(* IEC 61131-3 sources: Test-Git_ESME26/TestProgettoESME_26.fbsproj/TemplateFullProgrammingFramework_Migration.device.xml.v3^/Plc Logic.plclogic.xml.v3^/Application.application.xml.v3^/TemplateFullProgrammingFramework/EquipmentModules/SR_CharlyModule.pou.xml.v3^, 9 files *)

(* ---- Init_Reactions.act.st ---- *)
__METADATA__
{
  "v3Meta": {
    "objectGuid": "4aa47ba2-99d8-49fa-95b1-7f556ffac844",
    "objectTypeGuid": "8ac092e5-3128-4e26-9e7e-11016c6684f2",
    "embeddedObjectTypeGuids": [
      "3b83b776-fb25-43b8-99f2-3c507c9143fc"
    ],
    "properties": {},
    "subObjects": {}
  }
}

(* System generated code, only to be changed by experienced programmers *)
IF c_udiNumberOfSubModules < 1 THEN
	RETURN;
END_IF

(* Change of default reactions only on demand *)
(* Compare SR MainMachine Action Init_Reactions *)

xInitReactionsException := FALSE;

(*****************************************************************************************************************************************************)
(* Init ReactionTranslationMode *)

TPL.FC_InitReactionTranslationMode(	i_udiNumberOfSubModules			:= c_udiNumberOfSubModules,
									i_petReactionTranslationMode	:= ADR(aetReactionTranslationMode),
									q_etDiag						=> etDiag,
									q_etDiagExt						=> etDiagExtTPL);

IF etDiag <> GD.ET_Diag.Ok AND NOT xInitReactionsException THEN
	xInitReactionsException := TRUE;

	stInitReactionsException.sMsg := SE_CTBX.FC_MultiConcat(i_sString1 := 'InitReactionTranslationMode - ',
														i_sString2 := GD.FC_EtDiagToString(i_etDiag := etDiag),
														i_sString3 := ' - ',
														i_sString4 := TPL.FC_EtDiagExtToString(i_etDiagExt := etDiagExtTPL));
END_IF

(*****************************************************************************************************************************************************)
(* Init ReactionTranslationTable *)

TPL.FC_InitReactionTranslationTable(i_udiNumberOfSubModules			:= c_udiNumberOfSubModules,
									i_pstReactionTranslationTable	:= ADR(aastReactionTranslationTable),
									q_etDiag						=> etDiag,
									q_etDiagExt						=> etDiagExtTPL);

IF etDiag <> GD.ET_Diag.Ok AND NOT xInitReactionsException THEN
	xInitReactionsException := TRUE;

	stInitReactionsException.sMsg := SE_CTBX.FC_MultiConcat(i_sString1 := 'InitReactionTranslationTable - ',
														i_sString2 := GD.FC_EtDiagToString(i_etDiag := etDiag),
														i_sString3 := ' - ',
														i_sString4 := TPL.FC_EtDiagExtToString(i_etDiagExt := etDiagExtTPL));
END_IF

(*****************************************************************************************************************************************************)
(* Init ReactionTranslationJobs *)

TPL.FC_InitReactionTranslationJobs( i_udiNumberOfSubModules			:= c_udiNumberOfSubModules,
									i_pstReactionTranslationJobs	:= ADR(astReactionTranslationJobs),
									q_etDiag						=> etDiag,
									q_etDiagExt						=> etDiagExtTPL);

IF etDiag <> GD.ET_Diag.Ok AND NOT xInitReactionsException THEN
	xInitReactionsException := TRUE;

	stInitReactionsException.sMsg := SE_CTBX.FC_MultiConcat(i_sString1 := 'InitReactionTranslationJobs - ',
														i_sString2 := GD.FC_EtDiagToString(i_etDiag := etDiag),
														i_sString3 := ' - ',
														i_sString4 := TPL.FC_EtDiagExtToString(i_etDiagExt := etDiagExtTPL));
END_IF

(*****************************************************************************************************************************************************)
(* Set exception if any exception occurred *)

fbExceptionHandler.SetException(i_xExceptionActive	:= xInitReactionsException,
								iq_stException		:= stInitReactionsException,
								iq_stExceptionList	:= iq_stExceptionList);

xInitSuccessful := xInitSuccessful AND NOT xInitReactionsException;

etDiag := GD.ET_Diag.Ok;
(* End of system generated code, only to be changed by experienced programmers *)

(* ---- Init_Slave3.act.st ---- *)
__METADATA__
{
  "v3Meta": {
    "objectGuid": "d2282e85-0a4e-4bdb-8c08-0233ce9aa560",
    "objectTypeGuid": "8ac092e5-3128-4e26-9e7e-11016c6684f2",
    "embeddedObjectTypeGuids": [
      "3b83b776-fb25-43b8-99f2-3c507c9143fc"
    ],
    "properties": {},
    "subObjects": {}
  }
}

(* System generated code, could be modified for your application *)

(* Standard interface *)
astSubModuleInterface[c_udiSlave3].i_sModuleName := CONCAT(STR1 := iq_stStandardModuleItf.i_sModuleName, STR2 := ': Slave3');

astSubModuleInterface[c_udiSlave3].i_xLogEnable     := TRUE;
astSubModuleInterface[c_udiSlave3].i_wLogDataFilter := UDINT_TO_WORD(TPL.ET_LogDataFilter.ModuleDefault);

fbSlave3Module.RegisterLoggerPoint(i_ifParent := fbLoggerPoint, i_sName := 'Slave3', q_etDiag :=, q_etDiagExt :=);

(* AxisModule specific interface *)
stSlave3Interface.stMain.i_ifMaster 		:= i_ifMaster; (* Master *)
stSlave3Interface.stMain.i_ifDrive  		:= DRV_Slave3.Axis;
stSlave3Interface.stMain.iq_lencEncoder		:= LE_Slave3.Axis;
DRV_Slave3.Axis.SetErrorStopRamp(i_lrDeceleration := 50_000,
								  i_lrJerk		  := 500_000);

xDriveIsVirtual := FC_IsDriveVirtual(	i_ifDrive	:= stSlave3Interface.stMain.i_ifDrive,
										q_etDiag	=> etDiag,
										q_etDiagExt	=> etDiagExt,
										q_sMsg		=> sMsgBuffer);

IF etDiag <> GD.ET_Diag.Ok AND NOT xIsDriveVirtualException THEN
	stIsDriveVirtualException.etDiag 	:= etDiag;
	stIsDriveVirtualException.udiDiagExt:= etDiagExt;
	stIsDriveVirtualException.sDiagExt 	:= FC_EtDiagExtToString(i_etDiagExt := etDiagExt);
	stIsDriveVirtualException.sMsg 		:= sMsgBuffer;
	xIsDriveVirtualException 			:= TRUE;
END_IF

fbExceptionHandler.SetException(i_xExceptionActive	:= xIsDriveVirtualException,
								iq_stException		:= stIsDriveVirtualException,
								iq_stExceptionList	:= iq_stExceptionList);

xInitSuccessful := xInitSuccessful AND NOT xIsDriveVirtualException;
etDiag := GD.ET_Diag.Ok;

stSlave3Interface.stMain.i_lrMotionActiveVelLimit := 15.0; (* Limit for max. velocity of astAxisModuleInterface to switch output AxisMove in Units/s *)
stSlave3Interface.stMain.i_etMotionActiveVelType  := AXM_ET_MotionActiveVelType.RefVelocity;

stSlave3Interface.stMain.i_timMasterStop := T#1S;
stSlave3Interface.stMain.i_xHwLimitPos   := FALSE;
stSlave3Interface.stMain.i_xHwLimitNeg   := FALSE;

stSlave3Interface.stMain.stReducedVelocity.i_xEnableReducedVelocity		:= FALSE;
stSlave3Interface.stMain.stReducedVelocity.i_xOnlyLimitCheck			:= FALSE;
stSlave3Interface.stMain.stReducedVelocity.i_lrMaxReducedVelocity		:= 50.0;

stSlave3Interface.stMain.i_xStart := FALSE;

(***************************************************************************************************************************************************************************************************)
(*** Homing ***)
	IF xDriveIsVirtual THEN
		stSlave3Interface.stHome.i_etMode := PDL_ET_HomeMode.SetPosAxisAndLogEncoderPosition;			(* Homing Mode  in case of virtual axis *)
	ELSE
		stSlave3Interface.stHome.i_etMode := PDL_ET_HomeMode.PosDirectionPosEdgeSensor;						(* Homing Mode in case of real axis *)
	END_IF

	stSlave3Interface.stHome.i_xEnableInitAbsReadPos := FALSE;		(* TRUE : Restores the AxisPosition depending on the stHome.etMode
																			  If stHome.i_etMode is equal to PDL_ET_HomeMode.RestorePosFromAxisEncoder or
																			  to PDL_ET_HomeMode.WriteAxisEncoder, the encoder of the axis is read,
																			  or else the position will be restored from the retain area *)

 	stSlave3Interface.stHome.stSetpos.iq_pstRestorePosRetain := ADR(Grp_stRestorePositionAxis4);

	stSlave3Interface.stHome.i_xResetHomeOk := FALSE;

	(* Possible modes for homing mode Sensor:
		PDL_ET_HomeMode.PosDirectionPosEdgeSensor
		PDL_ET_HomeMode.NegDirectionPosEdgeSensor
		PDL_ET_HomeMode.NegDirectionNegEdgeSensor
		PDL_ET_HomeMode.PosDirectionNegEdgeSensor
	*)
	stSlave3Interface.stHome.stSensor.i_lrHomePosition			:= 0.0;			(* Position at the end of homing in units *)
	stSlave3Interface.stHome.stSensor.i_lrVel					:= 10.0;		(* Homing ceiling velocity in units/s *)
	stSlave3Interface.stHome.stSensor.i_lrAcc					:= 1000.0;		(* Homing acceleration in units/s^2 *)
	stSlave3Interface.stHome.stSensor.i_lrDec					:= 1000.0;		(* Homing deceleration in units/s^2 *)
	stSlave3Interface.stHome.stSensor.i_lrJerk					:= 10000.0;		(* Homing jerk in units/s^3 *)
	stSlave3Interface.stHome.stSensor.i_lrOffset				:= 0.0;			(* Offset from home signal in units *)
	stSlave3Interface.stHome.stSensor.i_lrMaxTravel				:= 720.0;		(* Max. travel for referencing by normal input *)
	stSlave3Interface.stHome.stSensor.i_xRotativeSystem			:= FALSE;		(* Rotative system true or false for referencing by normal input *)
	stSlave3Interface.stHome.stSensor.i_xSensor					:= FALSE;		(* Input for home signal. Can be a signal from a controller input. Has to be written cyclic. *)

	(* Possible Modes for homing mode LimitSwitch:
		PDL_ET_HomeMode.PosDirectionPosEdgeHWLimitPos		normally open contact / Closing contact
		PDL_ET_HomeMode.NegDirectionPosEdgeHWLimitNeg		normally open contact / Closing contact
		PDL_ET_HomeMode.NegDirectionNegEdgeHWLimitNeg		normally closed contact / Opening contact
		PDL_ET_HomeMode.PosDirectionNegEdgeHWLimitPos		normally closed contact / Opening contact
	*)
	stSlave3Interface.stHome.stLimitSwitch.i_lrHomePosition		:= 0.0;			(* Position at the end of homing in units *)
	stSlave3Interface.stHome.stLimitSwitch.i_lrVel				:= 10.0;		(* Homing ceiling velocity in units/s *)
	stSlave3Interface.stHome.stLimitSwitch.i_lrLowVel			:= 5.0;			(* Homing low ceiling velocity in units/s *)
	stSlave3Interface.stHome.stLimitSwitch.i_lrAcc				:= 1000.0;		(* Homing acceleration in units/s^2 *)
	stSlave3Interface.stHome.stLimitSwitch.i_lrDec				:= 1000.0;		(* Homing deceleration in units/s^2 *)
	stSlave3Interface.stHome.stLimitSwitch.i_lrJerk				:= 10000.0;		(* Homing jerk in units/s^3 *)
	stSlave3Interface.stHome.stLimitSwitch.i_lrOffset			:= 0.0;			(* Offset from home signal in units *)
	stSlave3Interface.stHome.stLimitSwitch.i_lrMaxTravel		:= 9999.0;		(* Max. travel for referencing normal input as a hardware limit *)

	(* Possible modes for homing mode MoveOnPos:
		PDL_ET_HomeMode.MoveOnPosAbs
	*)
	stSlave3Interface.stHome.stMoveOnPos.i_lrTarget				:= 0.0;			(* Position at the end of homing in units *)
	stSlave3Interface.stHome.stMoveOnPos.i_lrVel				:= 10.0;		(* Homing ceiling velocity in units/s *)
	stSlave3Interface.stHome.stMoveOnPos.i_lrAcc				:= 1000.0;		(* Homing acceleration in units/s^2 *)
	stSlave3Interface.stHome.stMoveOnPos.i_lrDec				:= 1000.0;		(* Homing deceleration in units/s^2 *)
	stSlave3Interface.stHome.stMoveOnPos.i_lrJerk				:= 10000.0;		(* Homing jerk in units/s^3 *)
	stSlave3Interface.stHome.stMoveOnPos.i_lrPeriod				:= 0.0;			(* Period of the axis *)
	stSlave3Interface.stHome.stMoveOnPos.i_xRotativeSystem		:= FALSE;		(* Rotative system true or false *)

	(* Possible modes for homing mode SetPos:
		PDL_ET_HomeMode.SetPosAxisPosition
		PDL_ET_HomeMode.SetPosLogEncoderPosition
		PDL_ET_HomeMode.SetPosAxisAndLogEncoderPosition
		PDL_ET_HomeMode.RestorePosFromAxisEncoder
		PDL_ET_HomeMode.RestorePosFromRetain
	*)
	stSlave3Interface.stHome.stSetpos.i_lrHomePosition			:= 0.0;			(* Position at the end of homing in units *)
	stSlave3Interface.stHome.stSetpos.i_lrEncoderPosition		:= 0.0;			(* Encoder position in units after homing *)
	stSlave3Interface.stHome.stSetpos.i_lrAbsEncOffset			:= 100.0;		(* Distance to the jump of axis encoder in units  *)
	stSlave3Interface.stHome.stSetpos.i_lrRestoreWindow			:= 180;			(* How far can the drive be away from is correct position *)
	stSlave3Interface.stHome.stSetpos.i_lrUserPeriod			:= 360;			(* Period of the axis *)
	stSlave3Interface.stHome.stSetPos.i_xKeepPowerDisabled 		:= FALSE;		(* Keep Power disabled during SetPosHoming true or false*)

	(* Possible modes for homing mode Torque:
		PDL_ET_HomeMode.PosDirectionMaxTorque
		PDL_ET_HomeMode.NegDirectionMaxTorque
	*)
	stSlave3Interface.stHome.stTorque.i_lrHomePosition			:= 0.0;			(* Position at the end of homing in units *)
	stSlave3Interface.stHome.stTorque.i_lrVel					:= 10.0;		(* Homing ceiling velocity in units/s *)
	stSlave3Interface.stHome.stTorque.i_lrAcc					:= 1000.0;		(* Homing acceleration in units/s^2 *)
	stSlave3Interface.stHome.stTorque.i_lrDec					:= 1000.0;		(* Homing deceleration in units/s^2 *)
	stSlave3Interface.stHome.stTorque.i_lrJerk					:= 10000.0;		(* Homing jerk in units/s^3 *)
	stSlave3Interface.stHome.stTorque.i_lrOffset				:= 0.0;			(* Offset from home signal in units *)
	stSlave3Interface.stHome.stTorque.i_lrMaxTravel				:= 9999.0;		(* Max. travel for referencing by torque *)
	stSlave3Interface.stHome.stTorque.i_lrMaxTorque				:= 0.0;			(* Torque for stop in Nm / referencing by torque *)
	stSlave3Interface.stHome.stTorque.i_diTorqueTime			:= 5;			(* Time in msec to hold torque *)

	(* Possible modes for homing mode TouchProbe:
		PDL_ET_HomeMode.PosDirectionPosEdgeTp
		PDL_ET_HomeMode.NegDirectionPosEdgeTp
		PDL_ET_HomeMode.NegDirectionNegEdgeTp
		PDL_ET_HomeMode.PosDirectionNegEdgeTp
	*)
	stSlave3Interface.stHome.stTouchProbe.i_lrHomePosition		:= 0.0;			(* Position at the end of homing in units *)
	stSlave3Interface.stHome.stTouchProbe.i_lrVel				:= 100.0;		(* Homing ceiling velocity in units/s *)
	stSlave3Interface.stHome.stTouchProbe.i_lrAcc				:= 1000.0;		(* Homing acceleration in units/s^2 *)
	stSlave3Interface.stHome.stTouchProbe.i_lrDec				:= 1000.0;		(* Homing deceleration in units/s^2 *)
	stSlave3Interface.stHome.stTouchProbe.i_lrJerk				:= 10000.0;		(* Homing jerk in units/s^3 *)
	stSlave3Interface.stHome.stTouchProbe.i_lrOffset			:= 30.0;		(* Offset from home signal in units *)
	stSlave3Interface.stHome.stTouchProbe.i_lrMaxTravel			:= 720.0;		(* Max. travel for referencing by TP *)
	stSlave3Interface.stHome.stTouchProbe.i_xRotativeSystem		:= TRUE;		(* Rotative system true or false for referencing by TP *)
 	stSlave3Interface.stHome.stTouchProbe.i_ifTouchProbe		:= 0;		(* Input for TP *)

	(* Possible modes for homing mode WritePos:
		PDL_ET_HomeMode.WriteAxisEncoder
	*)
	stSlave3Interface.stHome.stWritePos.i_lrHomePosition		:= 0.0;			(* Position at the end of homing in units *)
	stSlave3Interface.stHome.stWritePos.i_lrUserPeriod			:= 0.0;			(* Calculates Drive.Position into period ( units ) *)
	stSlave3Interface.stHome.stWritePos.i_lrAbsEncOffset		:= 100.0;		(* Distance to the jump of axis encoder in units *)

(***************************************************************************************************************************************************************************************************)
(*** Manual ***)
	stSlave3Interface.stManual.i_lrVel         := 50.0; (* Velocity in units/s *)
	stSlave3Interface.stManual.i_lrAcc         := 100.0; (* Acceleration in units/s^2 *)
	stSlave3Interface.stManual.i_lrDec         := 100.0; (* Deceleration in units/s^2 *)
	stSlave3Interface.stManual.i_lrJerk        := 1000.0; (* Jerk in units/s^3 *)
	stSlave3Interface.stManual.i_lrMaxDistance := 120.0; (* Max pathlengths for one step in units *)
	stSlave3Interface.stManual.i_xEndless      := FALSE; (* TRUE: jogging endless; Position between the periode; FALSE: jogging in steps. Position can be out of periode *)
	stSlave3Interface.stManual.i_lrPeriod      := 360.0; (* Period of the axis *)

(***************************************************************************************************************************************************************************************************)
(*** Cam ***)

	stSlave3Interface.stMultiCam.i_etCSModeSlave			:= PDL_ET_MultiCamCsModeSlave.SetSlavePositionToFirstCamPosition;		(* ColdStartMode Slave *)
	stSlave3Interface.stMultiCam.i_etCSModeMaster			:= PDL_ET_MultiCamCsModeMaster.SetMasterPositionToFirstCamPosition;		(* ColdStartMode Master *)
	stSlave3Interface.stMultiCam.i_etWSMode					:= PDL_ET_MultiCamWsMode.StoredCamMoveAlwaysNoPositionCheck;			(* WarmStartMode *)
	stSlave3Interface.stMultiCam.i_lrWSWindow				:= 5.0;											(* WarmStartWindow in Axis units *)
	stSlave3Interface.stMultiCam.i_lrWSVel					:= 10.0;										(* Velocity for WarmStart and CSModeSlave = PDL.ET_MultiCamCsModeSlave.MoveSlaveToFirstCamPosition in Units/s *)
	stSlave3Interface.stMultiCam.i_lrWSAcc					:= 1_000.0;										(* Acceleration and deceleration for Warmstart and CSModeSlave = PDL.ET_MultiCamCsModeSlave.MoveSlaveToFirstCamPosition in Units/s^2 *)
	stSlave3Interface.stMultiCam.i_lrWSJerk					:= 10_000.0;									(* Jerk for Warmstart and CSModeSlave = PDL.ET_MultiCamCsModeSlave.MoveSlaveToFirstCamPosition in units/s^3 *)
	stSlave3Interface.stMultiCam.i_diTXend					:= 2*G_diTaskIntervalInMs;	(* Time of XLowEnd and XHighEnd befor Xend or Xstart in msec*)
	stSlave3Interface.stMultiCam.i_lrInstantXLimMax			:= 180.0;											(* Switch off position at 'InstantNewCam' *)

	stSlave3Interface.stMultiCam.i_xEnableTabHandler		:= FALSE;										(* TRUE: TabHandler is enabled *)
	stSlave3Interface.stMultiCam.i_udiTableSelectNr			:= 0;							(* Number of table which is used in the next cycle *)

// 	stSlave3Interface.stMultiCam.i_xSetEncoderParameters	:= FALSE;										(* TRUE: The parameters MasterId, FeedConstand, GearIn and GearOut will be copyed into LEnc object *)
	stSlave3Interface.stMultiCam.i_xSetEncoderPosition		:= TRUE;										(* TRUE: Manipulation of LEnc object on startup OpMode MultiCam *)
	stSlave3Interface.stMultiCam.i_lrSetEncoderOffset		:= 0.0;											(* Master encoder offset *)
	stSlave3Interface.stMultiCam.i_xCheckEncoderPeriod		:= TRUE;										(* TRUE: Check of encoder period = 0. If encoder period <> 0 -> Exception *)

//	stSlave3Interface.stMultiCam.iq_xNewCam					:= FALSE;										(* TRUE: A new DataStruct will be load for next cycle. Will be reset when new cycle is started in case of stMultiCam.i_xEnableTabHandler = FALSE. *)
//	stSlave3Interface.stMultiCam.iq_xInstantNewCam			:= FALSE;										(* TRUE: A new DataStruct will be load. It will be active at master position stMultiCam.i_lrInstantXLimMax. Will be reset when ne DataStruct is active *)
//	stSlave3Interface.stMultiCam.iq_xChangeMaster			:= FALSE;										(* TRUE: Switch to a new Master. Will be reset when done. *)

// stSlave3Interface.stMultiCam.iq_stExt		;						(* Extended In of the Multicam FB, can be used if needed! *)

stSlave3Interface.stMultiCam.iq_astMotionPar[AXM_ET_ParId.User].diNumberOfCamPoints		:= 4;	(* DataStruct for the next cycle *)
stSlave3Interface.stMultiCam.iq_astMotionPar[AXM_ET_ParId.User].lrYPeriod				:= 0.0;

stSlave3Interface.stMultiCam.iq_astMotionPar[AXM_ET_ParId.User].astCamPoint[0].lrX		:= 0.0;
stSlave3Interface.stMultiCam.iq_astMotionPar[AXM_ET_ParId.User].astCamPoint[0].lrY		:= 0.0;
stSlave3Interface.stMultiCam.iq_astMotionPar[AXM_ET_ParId.User].astCamPoint[0].lrM		:= 0.0;
stSlave3Interface.stMultiCam.iq_astMotionPar[AXM_ET_ParId.User].astCamPoint[0].etCamType	:= PDL_ET_CamType.Poly5Com;
stSlave3Interface.stMultiCam.iq_astMotionPar[AXM_ET_ParId.User].astCamPoint[1].lrX		:= 60.0;
stSlave3Interface.stMultiCam.iq_astMotionPar[AXM_ET_ParId.User].astCamPoint[1].lrY		:= 30.0;
stSlave3Interface.stMultiCam.iq_astMotionPar[AXM_ET_ParId.User].astCamPoint[1].lrM		:= 1.0;
stSlave3Interface.stMultiCam.iq_astMotionPar[AXM_ET_ParId.User].astCamPoint[1].etCamType	:= PDL_ET_CamType.Straight;
stSlave3Interface.stMultiCam.iq_astMotionPar[AXM_ET_ParId.User].astCamPoint[2].lrX		:= 240.0;
stSlave3Interface.stMultiCam.iq_astMotionPar[AXM_ET_ParId.User].astCamPoint[2].lrY		:= 210.0;
stSlave3Interface.stMultiCam.iq_astMotionPar[AXM_ET_ParId.User].astCamPoint[2].lrM		:= 1.0;
stSlave3Interface.stMultiCam.iq_astMotionPar[AXM_ET_ParId.User].astCamPoint[2].etCamType	:= PDL_ET_CamType.Poly5Com;
stSlave3Interface.stMultiCam.iq_astMotionPar[AXM_ET_ParId.User].astCamPoint[3].lrX		:= 360.0;
stSlave3Interface.stMultiCam.iq_astMotionPar[AXM_ET_ParId.User].astCamPoint[3].lrY		:= 0.0;
stSlave3Interface.stMultiCam.iq_astMotionPar[AXM_ET_ParId.User].astCamPoint[3].lrM		:= 0.0;
stSlave3Interface.stMultiCam.iq_astMotionPar[AXM_ET_ParId.User].astCamPoint[3].etCamType	:= PDL_ET_CamType.Poly5Com;

stSlave3Interface.stMultiCam.iq_astMotionPar[AXM_ET_ParId.Idle].diUserTableId	:= UDINT_TO_DINT(AXM_ET_ParId.Idle);
stSlave3Interface.stMultiCam.iq_astMotionPar[AXM_ET_ParId.Start].diUserTableId	:= UDINT_TO_DINT(AXM_ET_ParId.Start);
stSlave3Interface.stMultiCam.iq_astMotionPar[AXM_ET_ParId.Cont].diUserTableId	:= UDINT_TO_DINT(AXM_ET_ParId.Cont);
stSlave3Interface.stMultiCam.iq_astMotionPar[AXM_ET_ParId.Stop].diUserTableId	:= UDINT_TO_DINT(AXM_ET_ParId.Stop);
stSlave3Interface.stMultiCam.iq_astMotionPar[AXM_ET_ParId.User].diUserTableId	:= UDINT_TO_DINT(AXM_ET_ParId.User);

(***************************************************************************************************************************************************************************************************)
(*** Endless ***)
	stSlave3Interface.stEndless.i_lrPeriod 					:= 500.0;		(* Period one cycle in units *)
	stSlave3Interface.stEndless.i_lrJerk 					:= 108000.0;	(* Jerk in units/s^3 *)
	stSlave3Interface.stEndless.i_lrStopPosition 			:= 120.0;		(* Stop position in units *)
	stSlave3Interface.stEndless.i_lrAcc  					:= 10800.0;		(* Acceleration in Units/s^2 *)
	stSlave3Interface.stEndless.i_lrDec  					:= 10800.0;		(* Deceleration in Units/s^2 *)
	stSlave3Interface.stEndless.i_lrVel 					:= 1080.0;   	(* Velocity in Units/s *)

(***************************************************************************************************************************************************************************************************)
(*** Pos ***)
	stSlave3Interface.stPos.i_etPosMode						:= PDL_ET_PosMode.Relative;		(* SYSTEMINTERFACE.ET_PosMode.Endless, SYSTEMINTERFACE.ET_PosMode.Relative, SYSTEMINTERFACE.ET_PosMode.Absolute *)
	stSlave3Interface.stPos.i_lrTarget 						:= 1440.0;		(* Target position or distance in Units *)
	stSlave3Interface.stPos.i_lrAcc 						:= 10800.0;		(* Acceleration in Units/s^2 *)
	stSlave3Interface.stPos.i_lrDec 						:= 10800.0;		(* Deceleration in Units/s^2 *)
	stSlave3Interface.stPos.i_lrJerk 						:= 108000.0;	(* Jerk in units/s^3 *)
	stSlave3Interface.stPos.i_lrVel 						:= 540.0;		(* Ceiling velocity in Units/s *)

// stSlave3Interface.stPos.i_xStop								:= FALSE;
(* End of system generated code, could be modified for your application *)

(* ---- Init_Slave4.act.st ---- *)
__METADATA__
{
  "v3Meta": {
    "objectGuid": "d38e3b28-2ba1-4cea-a02c-ff5eca86d734",
    "objectTypeGuid": "8ac092e5-3128-4e26-9e7e-11016c6684f2",
    "embeddedObjectTypeGuids": [
      "3b83b776-fb25-43b8-99f2-3c507c9143fc"
    ],
    "properties": {},
    "subObjects": {}
  }
}

(* System generated code, could be modified for your application *)

(* Standard interface *)
astSubModuleInterface[c_udiSlave4].i_sModuleName := CONCAT(STR1 := iq_stStandardModuleItf.i_sModuleName, STR2 := ': Slave4');

astSubModuleInterface[c_udiSlave4].i_xLogEnable     := TRUE;
astSubModuleInterface[c_udiSlave4].i_wLogDataFilter := UDINT_TO_WORD(TPL.ET_LogDataFilter.ModuleDefault);

fbSlave4Module.RegisterLoggerPoint(i_ifParent := fbLoggerPoint, i_sName := 'Slave4', q_etDiag :=, q_etDiagExt :=);

(* AxisModule specific interface *)
stSlave4Interface.stMain.i_ifMaster 		:= i_ifMaster; (* Master *)
stSlave4Interface.stMain.i_ifDrive  		:= DRV_Slave4.Axis;
stSlave4Interface.stMain.iq_lencEncoder		:= LE_Slave4.Axis;
DRV_Slave4.Axis.SetErrorStopRamp( i_lrDeceleration := 50_000,
								  i_lrJerk		   := 500_000);

xDriveIsVirtual := FC_IsDriveVirtual(	i_ifDrive	:= stSlave4Interface.stMain.i_ifDrive,
										q_etDiag	=> etDiag,
										q_etDiagExt	=> etDiagExt,
										q_sMsg		=> sMsgBuffer);

IF etDiag <> GD.ET_Diag.Ok AND NOT xIsDriveVirtualException THEN
	stIsDriveVirtualException.etDiag 	:= etDiag;
	stIsDriveVirtualException.udiDiagExt:= etDiagExt;
	stIsDriveVirtualException.sDiagExt 	:= FC_EtDiagExtToString(i_etDiagExt := etDiagExt);
	stIsDriveVirtualException.sMsg 		:= sMsgBuffer;
	xIsDriveVirtualException 			:= TRUE;
END_IF

fbExceptionHandler.SetException(i_xExceptionActive	:= xIsDriveVirtualException,
								iq_stException		:= stIsDriveVirtualException,
								iq_stExceptionList	:= iq_stExceptionList);

xInitSuccessful := xInitSuccessful AND NOT xIsDriveVirtualException;
etDiag := GD.ET_Diag.Ok;

stSlave4Interface.stMain.i_lrMotionActiveVelLimit := 15.0; (* Limit for max. velocity of astAxisModuleInterface to switch output AxisMove in Units/s *)
stSlave4Interface.stMain.i_etMotionActiveVelType  := AXM_ET_MotionActiveVelType.RefVelocity;

stSlave4Interface.stMain.i_timMasterStop := T#1S;
stSlave4Interface.stMain.i_xHwLimitPos   := FALSE;
stSlave4Interface.stMain.i_xHwLimitNeg   := FALSE;

stSlave4Interface.stMain.stReducedVelocity.i_xEnableReducedVelocity		:= FALSE;
stSlave4Interface.stMain.stReducedVelocity.i_xOnlyLimitCheck			:= FALSE;
stSlave4Interface.stMain.stReducedVelocity.i_lrMaxReducedVelocity		:= 50.0;

stSlave4Interface.stMain.i_xStart := FALSE;

(***************************************************************************************************************************************************************************************************)
(*** Homing ***)
	IF xDriveIsVirtual THEN
		stSlave4Interface.stHome.i_etMode := PDL_ET_HomeMode.SetPosAxisAndLogEncoderPosition;			(* Homing Mode  in case of virtual axis *)
	ELSE
		stSlave4Interface.stHome.i_etMode := PDL_ET_HomeMode.PosDirectionPosEdgeSensor;						(* Homing Mode in case of real axis *)
	END_IF

	stSlave4Interface.stHome.i_xEnableInitAbsReadPos := FALSE;		(* TRUE : Restores the AxisPosition depending on the stHome.etMode
																			  If stHome.i_etMode is equal to PDL_ET_HomeMode.RestorePosFromAxisEncoder or
																			  to PDL_ET_HomeMode.WriteAxisEncoder, the encoder of the axis is read,
																			  or else the position will be restored from the retain area *)

 	stSlave4Interface.stHome.stSetpos.iq_pstRestorePosRetain := ADR(Grp_stRestorePositionAxis5);

	stSlave4Interface.stHome.i_xResetHomeOk := FALSE;

	(* Possible modes for homing mode Sensor:
		PDL_ET_HomeMode.PosDirectionPosEdgeSensor
		PDL_ET_HomeMode.NegDirectionPosEdgeSensor
		PDL_ET_HomeMode.NegDirectionNegEdgeSensor
		PDL_ET_HomeMode.PosDirectionNegEdgeSensor
	*)
	stSlave4Interface.stHome.stSensor.i_lrHomePosition			:= 0.0;			(* Position at the end of homing in units *)
	stSlave4Interface.stHome.stSensor.i_lrVel					:= 10.0;		(* Homing ceiling velocity in units/s *)
	stSlave4Interface.stHome.stSensor.i_lrAcc					:= 1000.0;		(* Homing acceleration in units/s^2 *)
	stSlave4Interface.stHome.stSensor.i_lrDec					:= 1000.0;		(* Homing deceleration in units/s^2 *)
	stSlave4Interface.stHome.stSensor.i_lrJerk					:= 10000.0;		(* Homing jerk in units/s^3 *)
	stSlave4Interface.stHome.stSensor.i_lrOffset				:= 0.0;			(* Offset from home signal in units *)
	stSlave4Interface.stHome.stSensor.i_lrMaxTravel				:= 720.0;		(* Max. travel for referencing by normal input *)
	stSlave4Interface.stHome.stSensor.i_xRotativeSystem			:= FALSE;		(* Rotative system true or false for referencing by normal input *)
	stSlave4Interface.stHome.stSensor.i_xSensor					:= FALSE;		(* Input for home signal. Can be a signal from a controller input. Has to be written cyclic. *)

	(* Possible Modes for homing mode LimitSwitch:
		PDL_ET_HomeMode.PosDirectionPosEdgeHWLimitPos		normally open contact / Closing contact
		PDL_ET_HomeMode.NegDirectionPosEdgeHWLimitNeg		normally open contact / Closing contact
		PDL_ET_HomeMode.NegDirectionNegEdgeHWLimitNeg		normally closed contact / Opening contact
		PDL_ET_HomeMode.PosDirectionNegEdgeHWLimitPos		normally closed contact / Opening contact
	*)
	stSlave4Interface.stHome.stLimitSwitch.i_lrHomePosition		:= 0.0;			(* Position at the end of homing in units *)
	stSlave4Interface.stHome.stLimitSwitch.i_lrVel				:= 10.0;		(* Homing ceiling velocity in units/s *)
	stSlave4Interface.stHome.stLimitSwitch.i_lrLowVel			:= 5.0;			(* Homing low ceiling velocity in units/s *)
	stSlave4Interface.stHome.stLimitSwitch.i_lrAcc				:= 1000.0;		(* Homing acceleration in units/s^2 *)
	stSlave4Interface.stHome.stLimitSwitch.i_lrDec				:= 1000.0;		(* Homing deceleration in units/s^2 *)
	stSlave4Interface.stHome.stLimitSwitch.i_lrJerk				:= 10000.0;		(* Homing jerk in units/s^3 *)
	stSlave4Interface.stHome.stLimitSwitch.i_lrOffset			:= 0.0;			(* Offset from home signal in units *)
	stSlave4Interface.stHome.stLimitSwitch.i_lrMaxTravel		:= 9999.0;		(* Max. travel for referencing normal input as a hardware limit *)

	(* Possible modes for homing mode MoveOnPos:
		PDL_ET_HomeMode.MoveOnPosAbs
	*)
	stSlave4Interface.stHome.stMoveOnPos.i_lrTarget				:= 0.0;			(* Position at the end of homing in units *)
	stSlave4Interface.stHome.stMoveOnPos.i_lrVel				:= 10.0;		(* Homing ceiling velocity in units/s *)
	stSlave4Interface.stHome.stMoveOnPos.i_lrAcc				:= 1000.0;		(* Homing acceleration in units/s^2 *)
	stSlave4Interface.stHome.stMoveOnPos.i_lrDec				:= 1000.0;		(* Homing deceleration in units/s^2 *)
	stSlave4Interface.stHome.stMoveOnPos.i_lrJerk				:= 10000.0;		(* Homing jerk in units/s^3 *)
	stSlave4Interface.stHome.stMoveOnPos.i_lrPeriod				:= 0.0;			(* Period of the axis *)
	stSlave4Interface.stHome.stMoveOnPos.i_xRotativeSystem		:= FALSE;		(* Rotative system true or false *)

	(* Possible modes for homing mode SetPos:
		PDL_ET_HomeMode.SetPosAxisPosition
		PDL_ET_HomeMode.SetPosLogEncoderPosition
		PDL_ET_HomeMode.SetPosAxisAndLogEncoderPosition
		PDL_ET_HomeMode.RestorePosFromAxisEncoder
		PDL_ET_HomeMode.RestorePosFromRetain
	*)
	stSlave4Interface.stHome.stSetpos.i_lrHomePosition			:= 0.0;			(* Position at the end of homing in units *)
	stSlave4Interface.stHome.stSetpos.i_lrEncoderPosition		:= 0.0;			(* Encoder position in units after homing *)
	stSlave4Interface.stHome.stSetpos.i_lrAbsEncOffset			:= 100.0;		(* Distance to the jump of axis encoder in units  *)
	stSlave4Interface.stHome.stSetpos.i_lrRestoreWindow			:= 180;			(* How far can the drive be away from is correct position *)
	stSlave4Interface.stHome.stSetpos.i_lrUserPeriod			:= 360;			(* Period of the axis *)
	stSlave4Interface.stHome.stSetPos.i_xKeepPowerDisabled 		:= FALSE;		(* Keep Power disabled during SetPosHoming true or false*)

	(* Possible modes for homing mode Torque:
		PDL_ET_HomeMode.PosDirectionMaxTorque
		PDL_ET_HomeMode.NegDirectionMaxTorque
	*)
	stSlave4Interface.stHome.stTorque.i_lrHomePosition			:= 0.0;			(* Position at the end of homing in units *)
	stSlave4Interface.stHome.stTorque.i_lrVel					:= 10.0;		(* Homing ceiling velocity in units/s *)
	stSlave4Interface.stHome.stTorque.i_lrAcc					:= 1000.0;		(* Homing acceleration in units/s^2 *)
	stSlave4Interface.stHome.stTorque.i_lrDec					:= 1000.0;		(* Homing deceleration in units/s^2 *)
	stSlave4Interface.stHome.stTorque.i_lrJerk					:= 10000.0;		(* Homing jerk in units/s^3 *)
	stSlave4Interface.stHome.stTorque.i_lrOffset				:= 0.0;			(* Offset from home signal in units *)
	stSlave4Interface.stHome.stTorque.i_lrMaxTravel				:= 9999.0;		(* Max. travel for referencing by torque *)
	stSlave4Interface.stHome.stTorque.i_lrMaxTorque				:= 0.0;			(* Torque for stop in Nm / referencing by torque *)
	stSlave4Interface.stHome.stTorque.i_diTorqueTime			:= 5;			(* Time in msec to hold torque *)

	(* Possible modes for homing mode TouchProbe:
		PDL_ET_HomeMode.PosDirectionPosEdgeTp
		PDL_ET_HomeMode.NegDirectionPosEdgeTp
		PDL_ET_HomeMode.NegDirectionNegEdgeTp
		PDL_ET_HomeMode.PosDirectionNegEdgeTp
	*)
	stSlave4Interface.stHome.stTouchProbe.i_lrHomePosition		:= 0.0;			(* Position at the end of homing in units *)
	stSlave4Interface.stHome.stTouchProbe.i_lrVel				:= 100.0;		(* Homing ceiling velocity in units/s *)
	stSlave4Interface.stHome.stTouchProbe.i_lrAcc				:= 1000.0;		(* Homing acceleration in units/s^2 *)
	stSlave4Interface.stHome.stTouchProbe.i_lrDec				:= 1000.0;		(* Homing deceleration in units/s^2 *)
	stSlave4Interface.stHome.stTouchProbe.i_lrJerk				:= 10000.0;		(* Homing jerk in units/s^3 *)
	stSlave4Interface.stHome.stTouchProbe.i_lrOffset			:= 30.0;		(* Offset from home signal in units *)
	stSlave4Interface.stHome.stTouchProbe.i_lrMaxTravel			:= 720.0;		(* Max. travel for referencing by TP *)
	stSlave4Interface.stHome.stTouchProbe.i_xRotativeSystem		:= TRUE;		(* Rotative system true or false for referencing by TP *)
// 	stSlave4Interface.stHome.stTouchProbe.i_ifTouchProbe		:= TP_4;		(* Input for TP *)

	(* Possible modes for homing mode WritePos:
		PDL_ET_HomeMode.WriteAxisEncoder
	*)
	stSlave4Interface.stHome.stWritePos.i_lrHomePosition		:= 0.0;			(* Position at the end of homing in units *)
	stSlave4Interface.stHome.stWritePos.i_lrUserPeriod			:= 0.0;			(* Calculates Drive.Position into period ( units ) *)
	stSlave4Interface.stHome.stWritePos.i_lrAbsEncOffset		:= 100.0;		(* Distance to the jump of axis encoder in units *)

(***************************************************************************************************************************************************************************************************)
(*** Manual ***)
	stSlave4Interface.stManual.i_lrVel         := 50.0; (* Velocity in units/s *)
	stSlave4Interface.stManual.i_lrAcc         := 100.0; (* Acceleration in units/s^2 *)
	stSlave4Interface.stManual.i_lrDec         := 100.0; (* Deceleration in units/s^2 *)
	stSlave4Interface.stManual.i_lrJerk        := 1000.0; (* Jerk in units/s^3 *)
	stSlave4Interface.stManual.i_lrMaxDistance := 120.0; (* Max pathlengths for one step in units *)
	stSlave4Interface.stManual.i_xEndless      := FALSE; (* TRUE: jogging endless; Position between the periode; FALSE: jogging in steps. Position can be out of periode *)
	stSlave4Interface.stManual.i_lrPeriod      := 360.0; (* Period of the axis *)

(***************************************************************************************************************************************************************************************************)
(*** Cam ***)

	stSlave4Interface.stMultiCam.i_etCSModeSlave			:= PDL_ET_MultiCamCsModeSlave.SetSlavePositionToFirstCamPosition;		(* ColdStartMode Slave *)
	stSlave4Interface.stMultiCam.i_etCSModeMaster			:= PDL_ET_MultiCamCsModeMaster.SetMasterPositionToFirstCamPosition;		(* ColdStartMode Master *)
	stSlave4Interface.stMultiCam.i_etWSMode					:= PDL_ET_MultiCamWsMode.StoredCamMoveAlwaysNoPositionCheck;			(* WarmStartMode *)
	stSlave4Interface.stMultiCam.i_lrWSWindow				:= 5.0;											(* WarmStartWindow in Axis units *)
	stSlave4Interface.stMultiCam.i_lrWSVel					:= 10.0;										(* Velocity for WarmStart and CSModeSlave = PDL.ET_MultiCamCsModeSlave.MoveSlaveToFirstCamPosition in Units/s *)
	stSlave4Interface.stMultiCam.i_lrWSAcc					:= 1_000.0;										(* Acceleration and deceleration for Warmstart and CSModeSlave = PDL.ET_MultiCamCsModeSlave.MoveSlaveToFirstCamPosition in Units/s^2 *)
	stSlave4Interface.stMultiCam.i_lrWSJerk					:= 10_000.0;									(* Jerk for Warmstart and CSModeSlave = PDL.ET_MultiCamCsModeSlave.MoveSlaveToFirstCamPosition in units/s^3 *)
	stSlave4Interface.stMultiCam.i_diTXend					:= 2*G_diTaskIntervalInMs;	(* Time of XLowEnd and XHighEnd befor Xend or Xstart in msec*)
	stSlave4Interface.stMultiCam.i_lrInstantXLimMax			:= 180.0;											(* Switch off position at 'InstantNewCam' *)

	stSlave4Interface.stMultiCam.i_xEnableTabHandler		:= FALSE;										(* TRUE: TabHandler is enabled *)
	stSlave4Interface.stMultiCam.i_udiTableSelectNr			:= 0;							(* Number of table which is used in the next cycle *)

// 	stSlave4Interface.stMultiCam.i_xSetEncoderParameters	:= FALSE;										(* TRUE: The parameters MasterId, FeedConstand, GearIn and GearOut will be copyed into LEnc object *)
	stSlave4Interface.stMultiCam.i_xSetEncoderPosition		:= TRUE;										(* TRUE: Manipulation of LEnc object on startup OpMode MultiCam *)
	stSlave4Interface.stMultiCam.i_lrSetEncoderOffset		:= 0.0;											(* Master encoder offset *)
	stSlave4Interface.stMultiCam.i_xCheckEncoderPeriod		:= TRUE;										(* TRUE: Check of encoder period = 0. If encoder period <> 0 -> Exception *)

//	stSlave4Interface.stMultiCam.iq_xNewCam					:= FALSE;										(* TRUE: A new DataStruct will be load for next cycle. Will be reset when new cycle is started in case of stMultiCam.i_xEnableTabHandler = FALSE. *)
//	stSlave4Interface.stMultiCam.iq_xInstantNewCam			:= FALSE;										(* TRUE: A new DataStruct will be load. It will be active at master position stMultiCam.i_lrInstantXLimMax. Will be reset when ne DataStruct is active *)
//	stSlave4Interface.stMultiCam.iq_xChangeMaster			:= FALSE;										(* TRUE: Switch to a new Master. Will be reset when done. *)

// stSlave4Interface.stMultiCam.iq_stExt		;						(* Extended In of the Multicam FB, can be used if needed! *)

stSlave4Interface.stMultiCam.iq_astMotionPar[AXM_ET_ParId.User].diNumberOfCamPoints		:= 4;	(* DataStruct for the next cycle *)
stSlave4Interface.stMultiCam.iq_astMotionPar[AXM_ET_ParId.User].lrYPeriod				:= 0.0;

stSlave4Interface.stMultiCam.iq_astMotionPar[AXM_ET_ParId.User].astCamPoint[0].lrX		:= 0.0;
stSlave4Interface.stMultiCam.iq_astMotionPar[AXM_ET_ParId.User].astCamPoint[0].lrY		:= 0.0;
stSlave4Interface.stMultiCam.iq_astMotionPar[AXM_ET_ParId.User].astCamPoint[0].lrM		:= 0.0;
stSlave4Interface.stMultiCam.iq_astMotionPar[AXM_ET_ParId.User].astCamPoint[0].etCamType	:= PDL_ET_CamType.Poly5Com;
stSlave4Interface.stMultiCam.iq_astMotionPar[AXM_ET_ParId.User].astCamPoint[1].lrX		:= 60.0;
stSlave4Interface.stMultiCam.iq_astMotionPar[AXM_ET_ParId.User].astCamPoint[1].lrY		:= 30.0;
stSlave4Interface.stMultiCam.iq_astMotionPar[AXM_ET_ParId.User].astCamPoint[1].lrM		:= 1.0;
stSlave4Interface.stMultiCam.iq_astMotionPar[AXM_ET_ParId.User].astCamPoint[1].etCamType	:= PDL_ET_CamType.Straight;
stSlave4Interface.stMultiCam.iq_astMotionPar[AXM_ET_ParId.User].astCamPoint[2].lrX		:= 240.0;
stSlave4Interface.stMultiCam.iq_astMotionPar[AXM_ET_ParId.User].astCamPoint[2].lrY		:= 210.0;
stSlave4Interface.stMultiCam.iq_astMotionPar[AXM_ET_ParId.User].astCamPoint[2].lrM		:= 1.0;
stSlave4Interface.stMultiCam.iq_astMotionPar[AXM_ET_ParId.User].astCamPoint[2].etCamType	:= PDL_ET_CamType.Poly5Com;
stSlave4Interface.stMultiCam.iq_astMotionPar[AXM_ET_ParId.User].astCamPoint[3].lrX		:= 360.0;
stSlave4Interface.stMultiCam.iq_astMotionPar[AXM_ET_ParId.User].astCamPoint[3].lrY		:= 0.0;
stSlave4Interface.stMultiCam.iq_astMotionPar[AXM_ET_ParId.User].astCamPoint[3].lrM		:= 0.0;
stSlave4Interface.stMultiCam.iq_astMotionPar[AXM_ET_ParId.User].astCamPoint[3].etCamType	:= PDL_ET_CamType.Poly5Com;

stSlave4Interface.stMultiCam.iq_astMotionPar[AXM_ET_ParId.Idle].diUserTableId	:= UDINT_TO_DINT(AXM_ET_ParId.Idle);
stSlave4Interface.stMultiCam.iq_astMotionPar[AXM_ET_ParId.Start].diUserTableId	:= UDINT_TO_DINT(AXM_ET_ParId.Start);
stSlave4Interface.stMultiCam.iq_astMotionPar[AXM_ET_ParId.Cont].diUserTableId	:= UDINT_TO_DINT(AXM_ET_ParId.Cont);
stSlave4Interface.stMultiCam.iq_astMotionPar[AXM_ET_ParId.Stop].diUserTableId	:= UDINT_TO_DINT(AXM_ET_ParId.Stop);
stSlave4Interface.stMultiCam.iq_astMotionPar[AXM_ET_ParId.User].diUserTableId	:= UDINT_TO_DINT(AXM_ET_ParId.User);

(***************************************************************************************************************************************************************************************************)
(*** Endless ***)
	stSlave4Interface.stEndless.i_lrPeriod 					:= 500.0;		(* Period one cycle in units *)
	stSlave4Interface.stEndless.i_lrJerk 					:= 108000.0;	(* Jerk in units/s^3 *)
	stSlave4Interface.stEndless.i_lrStopPosition 			:= 120.0;		(* Stop position in units *)
	stSlave4Interface.stEndless.i_lrAcc  					:= 10800.0;		(* Acceleration in Units/s^2 *)
	stSlave4Interface.stEndless.i_lrDec  					:= 10800.0;		(* Deceleration in Units/s^2 *)
	stSlave4Interface.stEndless.i_lrVel 					:= 1080.0;   	(* Velocity in Units/s *)

(***************************************************************************************************************************************************************************************************)
(*** Pos ***)
	stSlave4Interface.stPos.i_etPosMode						:= PDL_ET_PosMode.Relative;		(* SYSTEMINTERFACE.ET_PosMode.Endless, SYSTEMINTERFACE.ET_PosMode.Relative, SYSTEMINTERFACE.ET_PosMode.Absolute *)
	stSlave4Interface.stPos.i_lrTarget 						:= 1440.0;		(* Target position or distance in Units *)
	stSlave4Interface.stPos.i_lrAcc 						:= 10800.0;		(* Acceleration in Units/s^2 *)
	stSlave4Interface.stPos.i_lrDec 						:= 10800.0;		(* Deceleration in Units/s^2 *)
	stSlave4Interface.stPos.i_lrJerk 						:= 108000.0;	(* Jerk in units/s^3 *)
	stSlave4Interface.stPos.i_lrVel 						:= 540.0;		(* Ceiling velocity in Units/s *)

// stSlave4Interface.stPos.i_xStop								:= FALSE;
(* End of system generated code, could be modified for your application *)

(* ---- Init_SubModules.act.st ---- *)
__METADATA__
{
  "v3Meta": {
    "objectGuid": "8e901039-7f2e-41e8-875d-6519455f0cb4",
    "objectTypeGuid": "8ac092e5-3128-4e26-9e7e-11016c6684f2",
    "embeddedObjectTypeGuids": [
      "3b83b776-fb25-43b8-99f2-3c507c9143fc"
    ],
    "properties": {},
    "subObjects": {}
  }
}

(* System generated code, could be modified for your application *)

(*** Module Group declaration ***)

aaudiSubModuleGroups[c_udiCharlyGroup1-TPL.GCL.Gc_udiGroupOffset,TPL.ET_Group.Member1] := 0;				(* There is no first element of the group c_diCharlyGroup1 *)
aaudiSubModuleGroups[c_udiCharlyGroup1-TPL.GCL.Gc_udiGroupOffset,TPL.ET_Group.Member2] := 0;				(* There is no second element of the group c_diCharlyGroup1 *)

aaudiSubModuleGroups[c_udiCharlyGroup2-TPL.GCL.Gc_udiGroupOffset,TPL.ET_Group.Member1] := c_udiSlave3;	(* The Slave3 is the first element of the group c_diCharlyGroup2 *)
aaudiSubModuleGroups[c_udiCharlyGroup2-TPL.GCL.Gc_udiGroupOffset,TPL.ET_Group.Member2] := c_udiSlave4;	(* The Slave4 is the second element of the group c_diCharlyGroup2 *)

(* End of system generated code, could be modified for your application *)

(* System generated code, do not change without consulting 'Schneider Electric Automation GmbH' - otherwise you risk instability!!!*)
xInitSubModulesException := FALSE;

(*****************************************************************************************************************************************************)
(* Set IDs of SubModules *)

TPL.FC_SetSubModuleIds(	i_udiMainModuleID			:= iq_stStandardModuleItf.i_udiModuleId,
						i_pstSubModulesItf			:= ADR(astSubModuleInterface),
						i_udiNumberOfSubModules		:= c_udiNumberOfSubModules,
						q_etDiag					=> etDiag,
						q_etDiagExt					=> etDiagExtTPL);

IF etDiag <> GD.ET_Diag.Ok AND NOT xInitSubModulesException THEN
	xInitSubModulesException := TRUE;

	stInitSubModulesException.sMsg := SE_CTBX.FC_MultiConcat(	i_sString1 := 'SetSubModuleIds - ',
															i_sString2 := GD.FC_EtDiagToString(i_etDiag := etDiag),
															i_sString3 := ' - ',
															i_sString4 := TPL.FC_EtDiagExtToString(i_etDiagExt := etDiagExtTPL));
END_IF

(*****************************************************************************************************************************************************)
(* Set exception if any exception occurred *)

fbExceptionHandler.SetException(i_xExceptionActive	:= xInitSubModulesException,
								iq_stException		:= stInitSubModulesException,
								iq_stExceptionList	:= iq_stExceptionList);

xInitSuccessful := xInitSuccessful AND NOT xInitSubModulesException;

etDiag := GD.ET_Diag.Ok;
(* End of system generated code, do not change without consulting 'Schneider Electric Automation GmbH' - otherwise you risk instability!!!*)

(* ---- Logic_Action.act.st ---- *)
__METADATA__
{
  "v3Meta": {
    "objectGuid": "4c63c3c9-7ae7-4f6a-8a63-3a1de13a49a1",
    "objectTypeGuid": "8ac092e5-3128-4e26-9e7e-11016c6684f2",
    "embeddedObjectTypeGuids": [
      "3b83b776-fb25-43b8-99f2-3c507c9143fc"
    ],
    "properties": {},
    "subObjects": {}
  }
}

(* This is an example of how to use the Positioning mode *)

IF stSlave4Interface.stMain.q_etOpMode = AXM_ET_OpMode.Positioning THEN
	IF stSlave4Interface.stMain.q_xMotionActive THEN
		(* There must be a rising edge at the xStart bit for initializing new Pos values, therefore it have to be reset. *)
		 stSlave4Interface.stMain.i_xStart := FALSE;
	END_IF

	CASE iPosState OF
		1: (* moving back *)
			(* Wait until the InPosition signal *)
			IF stSlave4Interface.stPos.q_xInPosition THEN
				(*Initialize new Pos values*)
				stSlave4Interface.stPos.i_lrTarget	:= -360.0;
				stSlave4Interface.stPos.i_etPosMode	:= PDL_ET_PosMode.Relative;

				IF fbLoggerPoint.etLogLevel >= APL.ET_LogLevel.StatusMessage THEN
					fbLoggerPoint.AddLogEntry(	i_etLogLevel	:= APL.ET_LogLevel.StatusMessage,
												i_etDiag		:= GD.ET_Diag.Ok,
												i_udiDiagExt	:= ET_DiagExt.Ok,
												i_sMessage		:= 'Logic: move axis in negative direction',
												q_etDiag		:= ,
												q_etDiagExt		:= );
				END_IF

				iPosState := 2;
			END_IF

		2: (* moving forward *)
			(* Wait until the InPosition signal *)
			IF stSlave4Interface.stPos.q_xInPosition THEN
				(* Initialize new Pos values *)
				stSlave4Interface.stPos.i_lrTarget	:= 360.0;
				stSlave4Interface.stPos.i_etPosMode	:= PDL_ET_PosMode.Relative;

				IF fbLoggerPoint.etLogLevel >= APL.ET_LogLevel.StatusMessage THEN
					fbLoggerPoint.AddLogEntry(	i_etLogLevel	:= APL.ET_LogLevel.StatusMessage,
												i_etDiag		:= GD.ET_Diag.Ok,
												i_udiDiagExt	:= ET_DiagExt.Ok,
												i_sMessage		:= 'Logic: move axis in positive direction',
												q_etDiag		:= ,
												q_etDiagExt		:= );
				END_IF

				iPosState := 1;
			END_IF
	END_CASE

	(* Start movement again and set new initialized values *)
	IF xFirstCall THEN
		xFirstCall := FALSE;

		stSlave4Interface.stMain.i_xStart := TRUE;

	ELSIF NOT stSlave4Interface.stMain.q_xMotionActive AND stSlave4Interface.stPos.q_xInPosition THEN
		stSlave4Interface.stMain.i_xStart := TRUE;
	END_IF
ELSE
	(* Set the SYSTEMINTERFACE.ET_PosMode.Absolute mode that the movement will start later at the last position. *)
	stSlave4Interface.stPos.i_etPosMode := PDL_ET_PosMode.Absolute;

	IF stSlave4Interface.stMain.q_etOpMode = AXM_ET_OpMode.Homing THEN
		(* Start with moving forward after homing *)
		stSlave4Interface.stPos.i_lrTarget := 360.0;

		iPosState := 1; (* next moving back *)
	END_IF
END_IF

(* ---- Output_Active.act.st ---- *)
__METADATA__
{
  "v3Meta": {
    "objectGuid": "05b7ecce-d158-4df2-a271-1322baec18fb",
    "objectTypeGuid": "8ac092e5-3128-4e26-9e7e-11016c6684f2",
    "embeddedObjectTypeGuids": [
      "3b83b776-fb25-43b8-99f2-3c507c9143fc"
    ],
    "properties": {},
    "subObjects": {}
  }
}

(* System generated code, only to be changed by experienced programmers *)
IF iq_stStandardModuleItf.q_udiSubModuleInException <> 0 THEN
	iq_stStandardModuleItf.q_etDiag		:= GD.ET_Diag.Ok;
	iq_stStandardModuleItf.q_udiDiagExt	:= ET_DiagExt.SubModuleInException;
	iq_stStandardModuleItf.q_sDiagExt		:= FC_EtDiagExtToString(i_etDiagExt := ET_DiagExt.SubModuleInException);
	iq_stStandardModuleItf.q_sMsg			:= '';
ELSE
	IF etDiagModuleController = GD.ET_Diag.Ok THEN
		iq_stStandardModuleItf.q_etDiag	:= etDiagModuleController;
		iq_stStandardModuleItf.q_sMsg		:= sMsgModuleController;

		CASE etDiagExtModuleController OF
			TPL.ET_DiagExt.DeactivatingSubModules :
				iq_stStandardModuleItf.q_udiDiagExt	:= ET_DiagExt.DeactivatingSubModules;
				iq_stStandardModuleItf.q_sDiagExt		:= FC_EtDiagExtToString(i_etDiagExt := ET_DiagExt.DeactivatingSubModules);
			TPL.ET_DiagExt.Disabled :
				iq_stStandardModuleItf.q_udiDiagExt	:= ET_DiagExt.Disabled;
				iq_stStandardModuleItf.q_sDiagExt		:= FC_EtDiagExtToString(i_etDiagExt := ET_DiagExt.Disabled);
			TPL.ET_DiagExt.ExecuteStep :
				iq_stStandardModuleItf.q_udiDiagExt	:= ET_DiagExt.ExecuteStep;
				iq_stStandardModuleItf.q_sDiagExt		:= FC_EtDiagExtToString(i_etDiagExt := ET_DiagExt.ExecuteStep);
			TPL.ET_DiagExt.Initializing :
				iq_stStandardModuleItf.q_udiDiagExt	:= ET_DiagExt.Initializing;
				iq_stStandardModuleItf.q_sDiagExt		:= FC_EtDiagExtToString(i_etDiagExt := ET_DiagExt.Initializing);
			TPL.ET_DiagExt.WaitAtNegativeStep :
				iq_stStandardModuleItf.q_udiDiagExt	:= ET_DiagExt.WaitAtNegativeStep;
				iq_stStandardModuleItf.q_sDiagExt		:= FC_EtDiagExtToString(i_etDiagExt := ET_DiagExt.WaitAtNegativeStep);
			TPL.ET_DiagExt.WaitCmdsDone :
				iq_stStandardModuleItf.q_udiDiagExt	:= ET_DiagExt.WaitCmdsDone;
				iq_stStandardModuleItf.q_sDiagExt		:= FC_EtDiagExtToString(i_etDiagExt := ET_DiagExt.WaitCmdsDone);
			TPL.ET_DiagExt.WaitForCmd :
				iq_stStandardModuleItf.q_udiDiagExt	:= ET_DiagExt.WaitForCmd;
				iq_stStandardModuleItf.q_sDiagExt		:= FC_EtDiagExtToString(i_etDiagExt := ET_DiagExt.WaitForCmd);
			ELSE
				iq_stStandardModuleItf.q_etDiag		:= GD. ET_Diag.UnexpectedProgramBehavior;
				iq_stStandardModuleItf.q_udiDiagExt	:= ET_DiagExt.UnknownStateModuleController;
				iq_stStandardModuleItf.q_sDiagExt		:= FC_EtDiagExtToString(i_etDiagExt := ET_DiagExt.UnknownStateModuleController);
		END_CASE
	ELSE
		iq_stStandardModuleItf.q_etDiag		:= GD.ET_Diag.DiagActive;
		iq_stStandardModuleItf.q_udiDiagExt	:= ET_DiagExt.ModuleControllerException;
		iq_stStandardModuleItf.q_sDiagExt		:= FC_EtDiagExtToString(i_etDiagExt := ET_DiagExt.ModuleControllerException);
		iq_stStandardModuleItf.q_sMsg			:= SE_CTBX.FC_MultiConcat(	i_sString1 := GD.FC_EtDiagToString(i_etDiag := etDiagModuleController),
																			i_sString2 := ' - ',
																			i_sString3 := TPL.FC_EtDiagExtToString(i_etDiagExt := etDiagExtModuleController),
																			i_sString4 := '');
	END_IF
END_IF

(* End of system generated code, only to be changed by experienced programmers *)

(* ---- RegisterLoggerPoint.meth.st ---- *)
METHOD RegisterLoggerPoint
VAR_INPUT
	i_ifParent	: APL.IF_LoggerPoint;
	i_sName		: STRING[80];
END_VAR
VAR_OUTPUT
	q_etDiag	: GD.ET_Diag := GD.ET_Diag.Ok;
	q_etDiagExt	: ET_DiagExt := ET_DiagExt.Ok;
END_VAR

fbLoggerPoint.RegisterLoggerPoint(	i_ifParent	:= i_ifParent,
									i_sName		:= i_sName,
									i_sType		:= 'Node Module',
									i_sSource	:= 'Program',
									q_etDiag	=> ,
									q_etDiagExt	=> );

(* ---- Start_Action.act.st ---- *)
__METADATA__
{
  "v3Meta": {
    "objectGuid": "5abc3db1-8b08-4e3a-9a94-3b606730b794",
    "objectTypeGuid": "8ac092e5-3128-4e26-9e7e-11016c6684f2",
    "embeddedObjectTypeGuids": [
      "3b83b776-fb25-43b8-99f2-3c507c9143fc"
    ],
    "properties": {},
    "subObjects": {}
  }
}

(* This step is active until the machine is being enabled *)

(* System generated code, do not change without consulting 'Schneider Electric Automation GmbH' - otherwise you risk instability!!! *)
iq_stStandardModuleItf.q_xActive			:= FALSE;
iq_stStandardModuleItf.q_xReady			:= FALSE;

iq_stStandardModuleItf.q_etDiag			:= GD.ET_Diag.Ok;
iq_stStandardModuleItf.q_udiDiagExt		:= ET_DiagExt.Disabled;
iq_stStandardModuleItf.q_sDiagExt			:= FC_EtDiagExtToString(i_etDiagExt := iq_stStandardModuleItf.q_udiDiagExt);
iq_stStandardModuleItf.q_sMsg				:= '';

iq_stStandardModuleItf.q_dwModuleType		:= TPL.ET_ModuleType.NodeModule;
iq_stStandardModuleItf.q_sModuleTypeName	:= 'NodeModule';
iq_stStandardModuleItf.q_udiModuleVersion	:= 1;
(* End of system generated code, do not change without consulting 'Schneider Electric Automation GmbH' - otherwise you risk instability!!! *)

(* System generated code, to be changed by experienced programmers *)
IF iq_stStandardModuleItf.iq_diCMD <> 0 AND NOT iq_stStandardModuleItf.i_xEnable THEN
	iq_stStandardModuleItf.iq_diCMD := 0;
END_IF
(* End of system generated code, to be changed by experienced programmers *)

(* Application specific code *)
(* ToDo: Add your application specific code here *)
;
(* End of application specific code *)

(* ---- UpdateStructs.act.st ---- *)
__METADATA__
{
  "v3Meta": {
    "objectGuid": "4b8e6845-be6c-47d0-9504-3441aa75f818",
    "objectTypeGuid": "8ac092e5-3128-4e26-9e7e-11016c6684f2",
    "embeddedObjectTypeGuids": [
      "3b83b776-fb25-43b8-99f2-3c507c9143fc"
    ],
    "properties": {},
    "subObjects": {}
  }
}

(* System generated code, do not change without consulting 'Schneider Electric Automation GmbH' - otherwise you risk instability!!!*)
fbDetectOnlineChange(	i_xEnable	:= TRUE,
						i_xDetect	:= TRUE,
						q_xActive	=> xDetectOnlineChangeActive,
						q_xReady	=> xDetectOnlineChangeReady,
						q_etDiag	=> etDetectOnlineChangeDiag,
						q_etDiagExt	=> etDetectOnlineChangeDiagExt,
						q_sMsg		=> sDetectOnlineChangeMsg,
						q_xChange	=> );

IF(NOT fbDetectOnlineChange.q_xChange) THEN
	RETURN;
END_IF

iq_stStandardModuleItf.iq_stExt.udiNumberOfSubModules 		:= c_udiNumberOfSubModules;
iq_stStandardModuleItf.iq_stExt.dwSubModulesItf		 		:= ADR(astSubModuleInterface);
iq_stStandardModuleItf.iq_stExt.pdwSubModulesAddItf 		:= ADR(adwSubModuleAddInterfaces);
iq_stStandardModuleItf.iq_stExt.pstListofCMDTables			:= ADR(astListOfCMDTables);
iq_stStandardModuleItf.iq_stExt.udiNumberOfCmdTables		:= c_udiNumberOfCMDTables;
(* End of system generated code, do not change without consulting 'Schneider Electric Automation GmbH' - otherwise you risk instability!!!*)

(* System generated code, could be modified for your application *)
xUpdateStructsException := FALSE;

(*****************************************************************************************************************************************************)
(* Update CmdTable - Prepare *)

TPL.FC_UpdateCmdTableListElement(	i_pstListofCMDTables	:= ADR(astListofCMDTables),
									i_udiNumberOfCmdTables	:= c_udiNumberOfCMDTables,
									i_diCMD					:= ET_Cmd.Prepare,
									i_pstCMDTable			:= ADR(astPrepareTable),
									q_etDiag				=> etDiag,
									q_etDiagExt				=> etDiagExtTPL);

IF etDiag <> GD.ET_Diag.Ok AND NOT xUpdateStructsException THEN
	xUpdateStructsException := TRUE;

	stUpdateStructsException.sMsg := SE_CTBX.FC_MultiConcat(i_sString1 := 'Update CmdTable: Prepare - ',
														i_sString2 := GD.FC_EtDiagToString(i_etDiag := etDiag),
														i_sString3 := ' - ',
														i_sString4 := TPL.FC_EtDiagExtToString(i_etDiagExt := etDiagExtTPL));
END_IF

(*****************************************************************************************************************************************************)
(* Update CmdTable - Auto *)

TPL.FC_UpdateCmdTableListElement(	i_pstListofCMDTables	:= ADR(astListofCMDTables),
									i_udiNumberOfCmdTables	:= c_udiNumberOfCMDTables,
									i_diCMD					:= ET_Cmd.Auto,
									i_pstCMDTable			:= ADR(astAutoTable),
									q_etDiag				=> etDiag,
									q_etDiagExt				=> etDiagExtTPL);

IF etDiag <> GD.ET_Diag.Ok AND NOT xUpdateStructsException THEN
	xUpdateStructsException := TRUE;

	stUpdateStructsException.sMsg := SE_CTBX.FC_MultiConcat(i_sString1 := 'Update CmdTable: Auto - ',
														i_sString2 := GD.FC_EtDiagToString(i_etDiag := etDiag),
														i_sString3 := ' - ',
														i_sString4 := TPL.FC_EtDiagExtToString(i_etDiagExt := etDiagExtTPL));
END_IF

(*****************************************************************************************************************************************************)
(* Update CmdTable - Manual *)

TPL.FC_UpdateCmdTableListElement(	i_pstListofCMDTables	:= ADR(astListofCMDTables),
									i_udiNumberOfCmdTables	:= c_udiNumberOfCMDTables,
									i_diCMD					:= ET_Cmd.Manual,
									i_pstCMDTable			:= ADR(astManualTable),
									q_etDiag				=> etDiag,
									q_etDiagExt				=> etDiagExtTPL);

IF etDiag <> GD.ET_Diag.Ok AND NOT xUpdateStructsException THEN
	xUpdateStructsException := TRUE;

	stUpdateStructsException.sMsg := SE_CTBX.FC_MultiConcat(i_sString1 := 'Update CmdTable: Manual - ',
														i_sString2 := GD.FC_EtDiagToString(i_etDiag := etDiag),
														i_sString3 := ' - ',
														i_sString4 := TPL.FC_EtDiagExtToString(i_etDiagExt := etDiagExtTPL));
END_IF

(*****************************************************************************************************************************************************)
(* Update CmdTable - Stop *)

TPL.FC_UpdateCmdTableListElement(	i_pstListofCMDTables	:= ADR(astListofCMDTables),
									i_udiNumberOfCmdTables	:= c_udiNumberOfCMDTables,
									i_diCMD					:= ET_Cmd.Stop,
									i_pstCMDTable			:= ADR(astStopTable),
									q_etDiag				=> etDiag,
									q_etDiagExt				=> etDiagExtTPL);

IF etDiag <> GD.ET_Diag.Ok AND NOT xUpdateStructsException THEN
	xUpdateStructsException := TRUE;

	stUpdateStructsException.sMsg := SE_CTBX.FC_MultiConcat(i_sString1 := 'Update CmdTable: Stop - ',
														i_sString2 := GD.FC_EtDiagToString(i_etDiag := etDiag),
														i_sString3 := ' - ',
														i_sString4 := TPL.FC_EtDiagExtToString(i_etDiagExt := etDiagExtTPL));
END_IF

(*****************************************************************************************************************************************************)
(* Update CmdTable - Start *)

TPL.FC_UpdateCmdTableListElement(	i_pstListofCMDTables	:= ADR(astListofCMDTables),
									i_udiNumberOfCmdTables	:= c_udiNumberOfCMDTables,
									i_diCMD					:= ET_Cmd.Start,
									i_pstCMDTable			:= ADR(astStartTable),
									q_etDiag				=> etDiag,
									q_etDiagExt				=> etDiagExtTPL);

IF etDiag <> GD.ET_Diag.Ok AND NOT xUpdateStructsException THEN
	xUpdateStructsException := TRUE;

	stUpdateStructsException.sMsg := SE_CTBX.FC_MultiConcat(i_sString1 := 'Update CmdTable: Start - ',
														i_sString2 := GD.FC_EtDiagToString(i_etDiag := etDiag),
														i_sString3 := ' - ',
														i_sString4 := TPL.FC_EtDiagExtToString(i_etDiagExt := etDiagExtTPL));
END_IF

(*****************************************************************************************************************************************************)
(* Update CmdTable - Abort *)

TPL.FC_UpdateCmdTableListElement(	i_pstListofCMDTables	:= ADR(astListofCMDTables),
									i_udiNumberOfCmdTables	:= c_udiNumberOfCMDTables,
									i_diCMD					:= ET_Cmd.Abort,
									i_pstCMDTable			:= ADR(astAbortTable),
									q_etDiag				=> etDiag,
									q_etDiagExt				=> etDiagExtTPL);

IF etDiag <> GD.ET_Diag.Ok AND NOT xUpdateStructsException THEN
	xUpdateStructsException := TRUE;

	stUpdateStructsException.sMsg := SE_CTBX.FC_MultiConcat(i_sString1 := 'Update CmdTable: Abort - ',
														i_sString2 := GD.FC_EtDiagToString(i_etDiag := etDiag),
														i_sString3 := ' - ',
														i_sString4 := TPL.FC_EtDiagExtToString(i_etDiagExt := etDiagExtTPL));
END_IF

(*****************************************************************************************************************************************************)
(* Update CmdTable - Hold *)

TPL.FC_UpdateCmdTableListElement(	i_pstListofCMDTables	:= ADR(astListofCMDTables),
									i_udiNumberOfCmdTables	:= c_udiNumberOfCMDTables,
									i_diCMD					:= ET_Cmd.Hold,
									i_pstCMDTable			:= ADR(astHoldTable),
									q_etDiag				=> etDiag,
									q_etDiagExt				=> etDiagExtTPL);

IF etDiag <> GD.ET_Diag.Ok AND NOT xUpdateStructsException THEN
	xUpdateStructsException := TRUE;

	stUpdateStructsException.sMsg := SE_CTBX.FC_MultiConcat(i_sString1 := 'Update CmdTable: Hold - ',
														i_sString2 := GD.FC_EtDiagToString(i_etDiag := etDiag),
														i_sString3 := ' - ',
														i_sString4 := TPL.FC_EtDiagExtToString(i_etDiagExt := etDiagExtTPL));
END_IF

(*****************************************************************************************************************************************************)
(* Update CmdTable - BrakeRelease *)

TPL.FC_UpdateCmdTableListElement(	i_pstListofCMDTables	:= ADR(astListofCMDTables),
									i_udiNumberOfCmdTables	:= c_udiNumberOfCMDTables,
									i_diCMD					:= ET_Cmd.BrakeRelease,
									i_pstCMDTable			:= ADR(astBrakeReleaseTable),
									q_etDiag				=> etDiag,
									q_etDiagExt				=> etDiagExtTPL);

IF etDiag <> GD.ET_Diag.Ok AND NOT xUpdateStructsException THEN
	xUpdateStructsException := TRUE;

	stUpdateStructsException.sMsg := SE_CTBX.FC_MultiConcat(i_sString1 := 'Update CmdTable: BrakeRelease - ',
														i_sString2 := GD.FC_EtDiagToString(i_etDiag := etDiag),
														i_sString3 := ' - ',
														i_sString4 := TPL.FC_EtDiagExtToString(i_etDiagExt := etDiagExtTPL));
END_IF

(*****************************************************************************************************************************************************)
(* Update AddInterface - Slave3 *)

AXM_FC_UpdateAddInterfaceStruct(	i_pdwSubModuleAddInterfaces	:= ADR(adwSubModuleAddInterfaces),
									i_udiSubModuleConstant		:= c_udiSlave3,
									iq_stAxisModuleItf			:= stSlave3Interface,
									q_etDiag					=> etDiag,
									q_etDiagExt					=> etDiagExtAXM);

IF etDiag <> GD.ET_Diag.Ok AND NOT xUpdateStructsException THEN
	xUpdateStructsException := TRUE;

	stUpdateStructsException.sMsg := SE_CTBX.FC_MultiConcat(i_sString1 := 'Update AddInterface: Slave3 - ',
														i_sString2 := GD.FC_EtDiagToString(i_etDiag := etDiag),
														i_sString3 := ' - ',
														i_sString4 := AXM_FC_EtDiagExtToString(i_etDiagExt := etDiagExtAXM));
END_IF

(*****************************************************************************************************************************************************)
(* Update AddInterface - Slave4 *)

AXM_FC_UpdateAddInterfaceStruct(	i_pdwSubModuleAddInterfaces	:= ADR(adwSubModuleAddInterfaces),
									i_udiSubModuleConstant		:= c_udiSlave4,
									iq_stAxisModuleItf			:= stSlave4Interface,
									q_etDiag					=> etDiag,
									q_etDiagExt					=> etDiagExtAXM);

IF etDiag <> GD.ET_Diag.Ok AND NOT xUpdateStructsException THEN
	xUpdateStructsException := TRUE;

	stUpdateStructsException.sMsg := SE_CTBX.FC_MultiConcat(i_sString1 := 'Update AddInterface: Slave4 - ',
														i_sString2 := GD.FC_EtDiagToString(i_etDiag := etDiag),
														i_sString3 := ' - ',
														i_sString4 := AXM_FC_EtDiagExtToString(i_etDiagExt := etDiagExtAXM));
END_IF

(*****************************************************************************************************************************************************)
(* Update AddInterface - Nocke1 *)

FC_UpdateExampleLeafModuleAddInterfaceStruct(	i_pdwSubModuleAddInterfaces		:= ADR(adwSubModuleAddInterfaces),
												i_udiSubModuleConstant			:= c_udiNocke1,
												iq_stExampleLeafModuleInterface	:= stNocke1Interface,
												q_etDiag						=> etDiag,
												q_etDiagExt						=> etDiagExtExampleLeaf);

IF etDiag <> GD.ET_Diag.Ok AND NOT xUpdateStructsException THEN
	xUpdateStructsException := TRUE;

	stUpdateStructsException.sMsg := SE_CTBX.FC_MultiConcat(i_sString1 := 'Update AddInterface: Nocke1 - ',
														i_sString2 := GD.FC_EtDiagToString(i_etDiag := etDiag),
														i_sString3 := ' - ',
														i_sString4 := FC_EtDiagExtExampleLeafModuleToString(i_etDiagExt := etDiagExtExampleLeaf));
END_IF

(*****************************************************************************************************************************************************)
(* Update ILS Data *)

// stSlave3Interface.stEndless.pstIlsData	:= ADR(G_stIlsData);
// stSlave3Interface.stMultiCam.pstIlsData	:= ADR(G_stIlsData);

// stSlave4Interface.stEndless.pstIlsData	:= ADR(G_stIlsData);
// stSlave4Interface.stMultiCam.pstIlsData	:= ADR(G_stIlsData);

(*****************************************************************************************************************************************************)
(* Set exception if any exception occurred *)

fbExceptionHandler.SetException(i_xExceptionActive	:= xUpdateStructsException,
								iq_stException		:= stUpdateStructsException,
								iq_stExceptionList	:= iq_stExceptionList);

xInitSuccessful := xInitSuccessful AND NOT xUpdateStructsException;

etDiag := GD.ET_Diag.Ok;
(* End of system generated code, could be modified for your application *)
